Fanuc KAREL source: KA00087.KL

PROGRAM KA00087
%NOLOCKGROUP
VAR
  SRC: JOINTPOS
  DST: BOOLEAN
BEGIN
  DST = SRC
END KA00087
